// FB_F_TRIG: 下降沿检测
// 描述: 检测TRUE到FALSE的跳变

FUNCTION_BLOCK FB_F_TRIG
VAR_INPUT
    IN  : BOOL;   // 待检测的布尔输入信号
END_VAR
VAR_OUTPUT
    Q   : BOOL;   // 下降沿检测输出 (一个周期内为TRUE)
END_VAR
VAR
    LastIN : BOOL := FALSE;
END_VAR

BEGIN
    // 检测下降沿: IN=FALSE且上一周期IN=TRUE
    #Q := NOT #IN AND #LastIN;
    #LastIN := #IN;

END_FUNCTION_BLOCK
